(* IEC 61131-3 sources: PLC-Static-Analysis/modules/plc-rules/src/test/resources/PLCA-Q015, 2 files *)

(* ---- compliant.st ---- *)
FUNCTION_BLOCK FB_Pump
VAR_INPUT
    bStart : BOOL;
    rSpeed : REAL;
    xEnable : BOOL;
    sName : STRING;
    tDelay : TIME;
    aValues : ARRAY[0..3] OF INT;
    pData : POINTER TO INT;
    eMode : E_Mode;
END_VAR
END_FUNCTION_BLOCK

TYPE E_Mode : (Off, On); END_TYPE

FUNCTION F_Add : INT
VAR_INPUT
    nA, nB : INT;
END_VAR
F_Add := nA + nB;
END_FUNCTION

(* ---- noncompliant.st ---- *)
FUNCTION_BLOCK Motor // PLCA-Q015
VAR_INPUT
    Start : BOOL; // PLCA-Q015
    speed : REAL; // PLCA-Q015
    nCount : INT;
    bigNumber : DINT; // PLCA-Q015
END_VAR
VAR
    timer : TON; // PLCA-Q015
    fbDelay : TON;
    stData : MotorData;
END_VAR
END_FUNCTION_BLOCK

TYPE MotorData : // PLCA-Q015
STRUCT
    bOk : BOOL;
END_STRUCT
END_TYPE

VAR_GLOBAL
    g_bReady : BOOL;
    gReady : BOOL; // PLCA-Q015
END_VAR
